PROGRAM main
  VAR
    S1 AT %IX0.0  : BOOL; (* marcha, NA *)
    S2 AT %IX0.1  : BOOL; (* paro, NC: TRUE sin pulsar *)
    KM1 AT %QX0.0 : BOOL; (* motor *)
    H1 AT %QX0.1  : BOOL; (* mantenimiento *)
    T_SEG         : TON;
    PULSO         : BOOL; (* TRUE una vuelta por segundo de marcha *)
    SEGUNDOS      : INT; (* horómetro: segundos de marcha *)
    HAY_TIEMPO    : BOOL; (* SEGUNDOS < 20 *)
  END_VAR
  VAR  (* added by the conversion: wires and edge detectors of the diagram *)
    _OR2_OUT : BOOL;
    _AND1_OUT : BOOL;
    _NOT10_OUT : BOOL;
    _AND8_OUT : BOOL;
    _ADD17_OUT : INT;
    _SEL14_OUT : INT;
    _GE21_OUT : BOOL;
  END_VAR

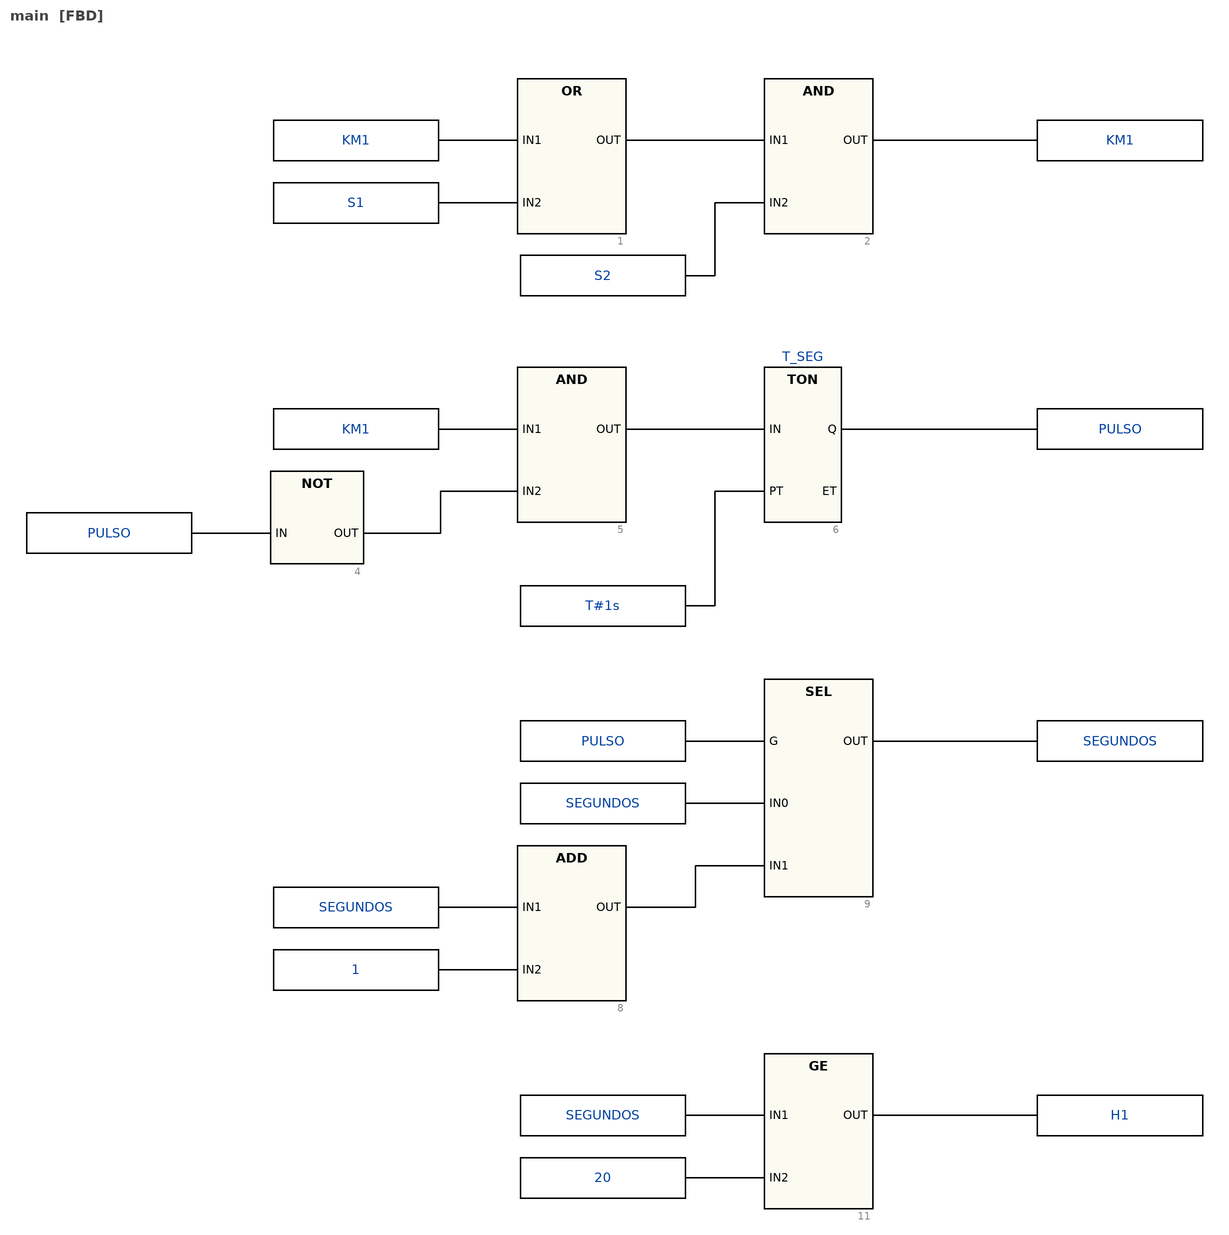
(* FBD diagram, written out as Structured Text *)
_OR2_OUT := KM1 OR S1;
_AND1_OUT := _OR2_OUT AND S2;
KM1 := _AND1_OUT;
_NOT10_OUT := NOT PULSO;
_AND8_OUT := KM1 AND _NOT10_OUT;
T_SEG(IN := _AND8_OUT, PT := T#1s);
PULSO := T_SEG.Q;
_ADD17_OUT := SEGUNDOS + 1;
_SEL14_OUT := SEL(PULSO, SEGUNDOS, _ADD17_OUT);
SEGUNDOS := _SEL14_OUT;
_GE21_OUT := SEGUNDOS >= 20;
H1 := _GE21_OUT;
END_PROGRAM
